// TIA Portal project "Project1" (V17)

(* hardware
DEVICE "S7-300/ET200M station_1"  S7-300 station
   slot 0: "Rail_0"  Rail  6ES7 390-1***0-0AA0
   slot 1: "PS 307 2A_1"  PS 307 2A  6ES7 307-1BA00-0AA0
   slot 2: "PLC_1"  CPU 315-2 PN/DP  6ES7 315-2EH14-0AB0  V3.2
      slot 2: "PROFINET interface_1"  PN-IO
         slot 1: "Port_1"  Port
         slot 2: "Port_2"  Port
   slot 3: "IM 365_1"  IM 365  6ES7 365-0BA01-0AA0
      slot 1: "IM send/receive interface_1"  6ES7 365-0BA00-0AA0
DEVICE "HMI_1"  TP1200 Comfort
   slot 0: "HMI_1"  TP1200 Comfort  6AV2 124-0MC01-0AX0  17.0.0.0
   slot 1: "HMI_RT_1"  TP1200 Comfort  6AV2 124-0MC01-0AX0  17.0.0.0
   slot 5: "HMI_1.IE_CP_1"  PROFINET Interface  17.0.0.0
      slot 1: "PROFINET Interface_1"  PROFINET Interface
         slot 1: "Port_1"  Port
         slot 2: "Port_2"  Port
   slot 7: "HMI_1.MPI/DP_CP_1"  MPI/DP Interface  17.0.0.0
*)

// ===== PLC "PLC_1"  CPU 315-2 PN/DP =====

VAR_GLOBAL   // PLC tag table "Default tag table"
   "START_BUTTON" AT %I0.3 : Bool;
   "STOP_BUTTON" AT %I0.4 : Bool;
   "MOTOR1" AT %Q0.0 : Bool;
   "MOTOR2" AT %Q0.1 : Bool;
   "MOTOR3" AT %Q0.2 : Bool;
   "SenRes1_LOW" AT %Q0.3 : Bool;
   "SenRes1_MID" AT %Q0.4 : Bool;
   "SenRes1_HIGH" AT %Q0.5 : Bool;
   "SenRes2_LOW" AT %Q0.6 : Bool;
   "SenRes2_MID" AT %Q0.7 : Bool;
   "SenRes2_HIGH" AT %Q1.0 : Bool;
   "SenFlow" AT %Q1.1 : Bool;
   "VALVE1" AT %Q1.2 : Bool;
   "VALVE2" AT %Q1.3 : Bool;
   "SYS_STATE" AT %Q1.4 : Bool;
   "M1_WORK_2S" AT %Q1.5 : Bool;
   "M2_DWORK_2S" AT %Q1.6 : Bool;
   "MID_DRAIN" AT %Q1.7 : Bool;
   "FILLED" AT %Q2.0 : Bool;
END_VAR

ORGANIZATION_BLOCK "Main"   // OB1, LAD
TITLE = "Main Program Sweep (Cycle)"
{ S7_Optimized_Access := 'FALSE' }
VERSION : 0.1
   VAR_TEMP
      OB1_EV_CLASS : Byte;   // Bits 0-3 = 1 (Coming event), Bits 4-7 = 1 (Event class 1)
      OB1_SCAN_1 : Byte;   // 1 (Cold restart scan 1 of OB 1), 3 (Scan 2-n of OB 1)
      OB1_PRIORITY : Byte;   // Priority of OB Execution
      OB1_OB_NUMBR : Byte;   // 1 (Organization block 1, OB1)
      OB1_RESERVED_1 : Byte;   // Reserved for system
      OB1_RESERVED_2 : Byte;   // Reserved for system
      OB1_PREV_CYCLE : Int;   // Cycle time of previous OB1 scan (milliseconds)
      OB1_MIN_CYCLE : Int;   // Minimum cycle time of OB1 (milliseconds)
      OB1_MAX_CYCLE : Int;   // Maximum cycle time of OB1 (milliseconds)
      OB1_DATE_TIME : Date_And_Time;   // Date and time OB1 started
   END_VAR
BEGIN

REGION Network 1
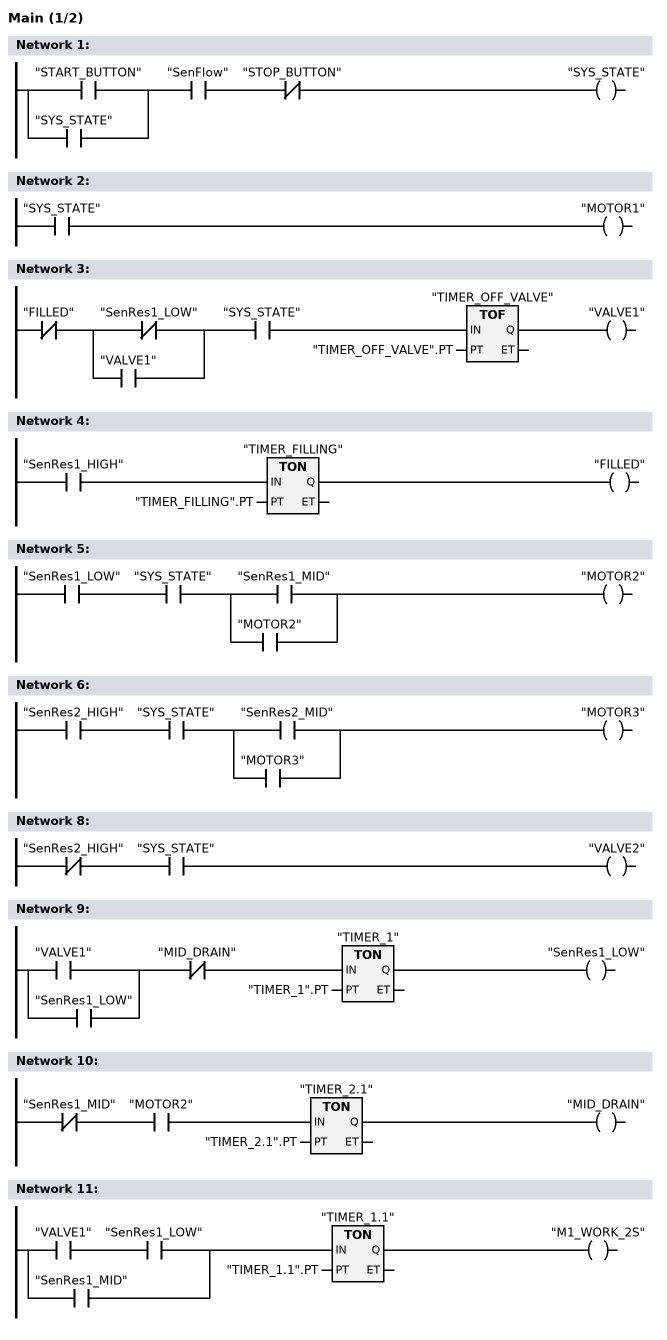
   RUNG wire#powerrail
      Contact( "START_BUTTON" )
      wire#w1
      Contact( "SenFlow" )
      I_Contact( "STOP_BUTTON" )
      Coil( "SYS_STATE" )
   END_RUNG
   RUNG wire#powerrail
      Contact( "SYS_STATE" )
   END_RUNG wire#w1
   // the same network as SCL:
   "SYS_STATE" := ("START_BUTTON" OR "SYS_STATE") AND "SenFlow" AND NOT "STOP_BUTTON";
END_REGION

REGION Network 2
   RUNG wire#powerrail
      Contact( "SYS_STATE" )
      Coil( "MOTOR1" )
   END_RUNG
   // the same network as SCL:
   "MOTOR1" := "SYS_STATE";
END_REGION

REGION Network 3
   "TIMER_OFF_VALVE".TOF(IN := NOT "FILLED" AND (NOT "SenRes1_LOW" OR "VALVE1") AND "SYS_STATE",
                         PT := "TIMER_OFF_VALVE".PT);
   "VALVE1" := "TIMER_OFF_VALVE".Q;
END_REGION

REGION Network 4
   "TIMER_FILLING".TON(IN := "SenRes1_HIGH", PT := "TIMER_FILLING".PT);
   "FILLED" := "TIMER_FILLING".Q;
END_REGION

REGION Network 5
   RUNG wire#powerrail
      Contact( "SenRes1_LOW" )
      Contact( "SYS_STATE" )
      wire#w1
      Contact( "SenRes1_MID" )
      wire#w2
      Coil( "MOTOR2" )
   END_RUNG
   RUNG wire#w1
      Contact( "MOTOR2" )
   END_RUNG wire#w2
   // the same network as SCL:
   "MOTOR2" := "SenRes1_LOW" AND "SYS_STATE" AND ("SenRes1_MID" OR "MOTOR2");
END_REGION

REGION Network 6
   RUNG wire#powerrail
      Contact( "SenRes2_HIGH" )
      Contact( "SYS_STATE" )
      wire#w1
      Contact( "SenRes2_MID" )
      wire#w2
      Coil( "MOTOR3" )
   END_RUNG
   RUNG wire#w1
      Contact( "MOTOR3" )
   END_RUNG wire#w2
   // the same network as SCL:
   "MOTOR3" := "SenRes2_HIGH" AND "SYS_STATE" AND ("SenRes2_MID" OR "MOTOR3");
END_REGION

REGION Network 8
   RUNG wire#powerrail
      I_Contact( "SenRes2_HIGH" )
      Contact( "SYS_STATE" )
      Coil( "VALVE2" )
   END_RUNG
   // the same network as SCL:
   "VALVE2" := NOT "SenRes2_HIGH" AND "SYS_STATE";
END_REGION

REGION Network 9
   "TIMER_1".TON(IN := ("VALVE1" OR "SenRes1_LOW") AND NOT "MID_DRAIN", PT := "TIMER_1".PT);
   "SenRes1_LOW" := "TIMER_1".Q;
END_REGION

REGION Network 10
   "TIMER_2.1".TON(IN := NOT "SenRes1_MID" AND "MOTOR2", PT := "TIMER_2.1".PT);
   "MID_DRAIN" := "TIMER_2.1".Q;
END_REGION

REGION Network 11
   "TIMER_1.1".TON(IN := ("VALVE1" AND "SenRes1_LOW") OR "SenRes1_MID", PT := "TIMER_1.1".PT);
   "M1_WORK_2S" := "TIMER_1.1".Q;
END_REGION

REGION Network 12
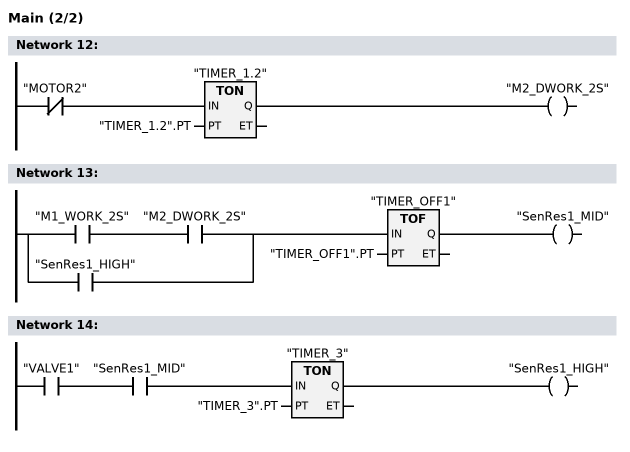
   "TIMER_1.2".TON(IN := NOT "MOTOR2", PT := "TIMER_1.2".PT);
   "M2_DWORK_2S" := "TIMER_1.2".Q;
END_REGION

REGION Network 13
   "TIMER_OFF1".TOF(IN := ("M1_WORK_2S" AND "M2_DWORK_2S") OR "SenRes1_HIGH", PT := "TIMER_OFF1".PT);
   "SenRes1_MID" := "TIMER_OFF1".Q;
END_REGION

REGION Network 14
   "TIMER_3".TON(IN := "VALVE1" AND "SenRes1_MID", PT := "TIMER_3".PT);
   "SenRes1_HIGH" := "TIMER_3".Q;
END_REGION
END_ORGANIZATION_BLOCK

(* ===== HMI "HMI_RT_1" =====
system functions are stored by id; their names below are inferred from use
connection "HMI_Connection_1": ETHERNET, SIMATIC S7 300/400 MPI

HMI tags "Default tag table"
   "START_BUTTON" : Bool = PLC START_BUTTON AT %I0.3, 1 s
   "STOP_BUTTON" : Bool = PLC STOP_BUTTON AT %I0.4, 1 s
   "SYS_STATE" : Bool = PLC SYS_STATE AT %Q1.4, 1 s
   "SenRes1_HIGH" : Bool = PLC SenRes1_HIGH AT %Q0.5, 1 s
   "SenRes2_LOW" : Bool = PLC SenRes2_LOW AT %Q0.6, 1 s
   "SenRes1_LOW" : Bool = PLC SenRes1_LOW AT %Q0.3, 1 s
   "VALVE1" : Bool = PLC VALVE1 AT %Q1.2, 1 s
   "VALVE2" : Bool = PLC VALVE2 AT %Q1.3, 1 s
   "SenFlow" : Bool = PLC SenFlow AT %Q1.1, 1 s
   "Tag_ScreenNumber" : UInt, internal
   "SenRes1_MID" : Bool = PLC SenRes1_MID AT %Q0.4, 1 s
   "MOTOR1" : Bool = PLC MOTOR1 AT %Q0.0, 1 s
   "MOTOR2" : Bool = PLC MOTOR2 AT %Q0.1, 1 s
   "MOTOR3" : Bool = PLC MOTOR3 AT %Q0.2, 1 s
   "SenRes2_MID" : Bool = PLC SenRes2_MID AT %Q0.7, 1 s
   "SenRes2_HIGH" : Bool = PLC SenRes2_HIGH AT %Q1.0, 1 s

screen "Root screen" 1280x757, template "Template_1"
   on GenerateScreen: SetTag("Tag_ScreenNumber", 1)
   SymbolLibrary "Symbol library_26" at 622,81 size 131x30
   SymbolLibrary "Symbol library_7" at 180,109 size 33x309
      Appearance <- "SYS_STATE"
   SymbolLibrary "Symbol library_25" at 211,79 size 175x30
      Appearance <- "SYS_STATE"
   SymbolLibrary "Symbol library_10" at 413,340 size 33x91
   Button "Button_1" at 18,81 size 146x67; TextOff 'Start'
      on Click: SetBit("START_BUTTON"); ResetBit("STOP_BUTTON")
   SymbolLibrary "Symbol library_3" at 394,418 size 86x118
      Appearance <- "MOTOR2"
   SymbolLibrary "Symbol library_5" at 778,336 size 33x91
   SymbolLibrary "Symbol library_1" at 699,42 size 189x318
   SymbolLibrary "Symbol library_11" at 755,414 size 86x118
      Appearance <- "MOTOR3"
   SymbolLibrary "Symbol library_14" at 834,422 size 131x30
   SymbolLibrary "Symbol library_15" at 474,429 size 85x30
   SymbolLibrary "Symbol library_9" at 181,69 size 60x53
      Appearance <- "SYS_STATE"
   SymbolLibrary "Symbol library_6" at 960,172 size 313x333
   SymbolLibrary "Symbol library_2" at 335,44 size 189x316
   SymbolLibrary "Symbol library_24" at 242,17 size 85x91
      Appearance <- "VALVE1"
      ProcessValue <- "VALVE1"
   SymbolLibrary "Symbol library_27" at 164,14 size 63x54
      Appearance <- "SYS_STATE"
   SymbolLibrary "Symbol library_29" at 148,391 size 65x60
      Appearance <- "SenFlow"
   Button "Button_2" at 18,163 size 146x67; TextOff 'Stop'
      on Click: SetBit("STOP_BUTTON"); ResetBit("START_BUTTON")
   Button "Button_3" at 39,539 size 194x60; TextOff 'Man Stop 1'
      on Click: SetBit("STOP_BUTTON")
   Button "Button_4" at 349,539 size 189x60; TextOff 'Man Stop 2'
      on Click: SetBit("STOP_BUTTON")
   Button "Button_5" at 696,539 size 196x60; TextOff 'Man Stop 3'
      on Click: SetBit("STOP_BUTTON")
   Circle "Circle_1" at 976,40 size 111x111
      Appearance <- "SYS_STATE"
   Circle "Circle_2" at 1118,42 size 111x111
      Appearance <- "SYS_STATE"
   Circle "Circle_5" at 319,476 size 53x53
      Appearance <- "MOTOR2"
   Circle "Circle_6" at 318,416 size 53x53
      Appearance <- "MOTOR2"
   Circle "Circle_3" at 19,476 size 53x53
      Appearance <- "MOTOR1"
   Circle "Circle_4" at 18,416 size 53x53
      Appearance <- "MOTOR1"
   Circle "Circle_7" at 684,476 size 53x53
      Appearance <- "MOTOR3"
   Circle "Circle_8" at 683,416 size 53x53
      Appearance <- "MOTOR3"
   SymbolLibrary "Symbol library_4" at 83,415 size 86x118
      Appearance <- "MOTOR1"
   SymbolLibrary "Symbol library_16" at 568,70 size 63x53
   SymbolLibrary "Symbol library_28" at 626,19 size 70x90
      ProcessValue <- "VALVE2"
      Appearance <- "VALVE2"
   SymbolLibrary "Symbol library_30" at 553,16 size 63x54
   SymbolLibrary "Symbol library_12" at 535,399 size 65x60
   SymbolLibrary "Symbol library_13" at 567,123 size 33x277
   Polygon "Polygon_3" at 366,274 size 122x79
      Visibility <- "SenRes1_LOW"
   Polygon "Polygon_4" at 729,276 size 122x79
      Visibility <- "SenRes2_LOW"
   Polygon "Polygon_5" at 338,171 size 181x98
      Visibility <- "SenRes1_MID"
   SymbolLibrary "Symbol library_18" at 492,244 size 65x27
      Appearance <- "SenRes1_LOW"
   Polygon "Polygon_6" at 337,61 size 184x111
      Visibility <- "SenRes1_HIGH"
   SymbolLibrary "Symbol library_20" at 492,54 size 65x27
      Appearance <- "SenRes1_HIGH"
   SymbolLibrary "Symbol library_19" at 492,161 size 65x27
      Appearance <- "SenRes1_MID"
   SymbolLibrary "Symbol library_8" at 154,336 size 67x70
      Appearance <- "SenFlow"
   Polygon "Polygon_1" at 355,264 size 149x90
      Visibility <- "SenRes1_LOW"
   Polygon "Polygon_2" at 720,261 size 145x94
      Visibility <- "SenRes2_LOW"
   Polygon "Polygon_8" at 702,169 size 181x98
      Visibility <- "SenRes2_MID"
   SymbolLibrary "Symbol library_21" at 861,244 size 65x27
      Appearance <- "SenRes2_LOW"
   Polygon "Polygon_9" at 699,59 size 184x111
      Visibility <- "SenRes2_HIGH"
   SymbolLibrary "Symbol library_22" at 861,161 size 65x27
      Appearance <- "SenRes2_MID"
   SymbolLibrary "Symbol library_23" at 861,54 size 65x27
      Appearance <- "SenRes2_HIGH"
   Button "Button_6" at 14,342 size 126x51; TextOff 'FLUX ON/OFF'
      on Click: InvertBit("SenFlow")

Template "Template_1" 1280x757
   Button "Exit" at 1840,960 size 78x58; TextOff 'Exit'; PictureOff "ExitRuntime_TP2200_Comfort_V2_TR"; PictureOn "ExitRuntime_TP2200_Comfort_V2_TR"
      on Release: StopRuntime(0)
   Button "Template_Button" at 1760,960 size 78x58; TextOff 'Text'
   Button "Template_Button_1" at 1680,960 size 78x58; TextOff 'Text'
   Button "Template_Button_2" at 1600,960 size 78x58; TextOff 'Text'
   Button "Template_Button_3" at 1520,960 size 78x58; TextOff 'Text'
   Button "Template_Button_4" at 1440,960 size 78x58; TextOff 'Text'
   Button "Template_Button_5" at 1360,960 size 78x58; TextOff 'Text'
   Button "Template_Button_6" at 1280,960 size 78x58; TextOff 'Text'
   Button "Template_Button_7" at 1200,960 size 78x58; TextOff 'Text'
   Button "Template_Button_8" at 1120,960 size 78x58; TextOff 'Text'
   Button "Template_Button_9" at 1040,960 size 78x58; TextOff 'Text'
   Button "Template_Button_10" at 960,960 size 78x58; TextOff 'Text'
   Button "Template_Button_11" at 881,960 size 78x58; TextOff 'Text'
   Button "Template_Button_12" at 801,960 size 78x58; TextOff 'Text'
   Button "Template_Button_13" at 721,960 size 78x58; TextOff 'Text'
   Button "Template_Button_14" at 641,960 size 78x58; TextOff 'Text'
   Button "Template_Button_15" at 561,960 size 78x58; TextOff 'Text'
   Button "Template_Button_16" at 481,960 size 78x58; TextOff 'Text'
   Button "Template_Button_17" at 401,960 size 78x58; TextOff 'Text'
   Button "Template_Button_18" at 321,960 size 78x58; TextOff 'Text'
   Button "Template_Button_19" at 241,960 size 78x58; TextOff 'Text'
   Button "Template_Button_20" at 161,960 size 78x58; TextOff 'Text'
   Button "Template_Button_21" at 81,960 size 78x58; TextOff 'Text'
   Button "Start screen" at 1,960 size 78x58; TextOff 'Start screen'; PictureOff "NavigateHome_TP2200_Comfort_V2_TR"; PictureOn "NavigateHome_TP2200_Comfort_V2_TR"
      on Release: ActivateScreen("Root screen", 0)

VB script "VBFunction_1"
   'Tip:
   ' 1. Use the <CTRL+SPACE> or <CTRL+I> shortcut to open a list of all objects and functions
   ' 2. Write the code using the HMI Runtime object.
   '  Example: HmiRuntime.Screens("Screen_1").
   ' 3. Use the <CTRL+J> shortcut to create an object reference.
   'Write the code as of this position:
*)